(* IEC 61131-3 sources: codesys-ai-industrial-robot-control/plc/src/Comm, 4 files *)

(* ---- GVL_Bridge.st ---- *)
// Exchange with the Python bridge over OPC UA (published by the symbol configuration).
// Tag names for the bridge: config/opcua_tags.yaml. In Phase 1, tests write the inputs.
{attribute 'qualified_only'}
{attribute 'symbol' := 'readwrite'}
VAR_GLOBAL
    // --- inputs (bridge -> PLC) ---
    xHeartbeat : BOOL;                                     // toggled by the bridge every cycle
    xTwinActive : BOOL;                                    // the twin delivers joint feedback
    aJointPosFb : ARRAY[1..6] OF LREAL;                    // measured joint positions [deg]
    aJointTorqueFb : ARRAY[1..6] OF LREAL;                 // measured joint torques [Nm]
    udiFeedbackSeq : UDINT;                                // increments with every feedback sample
    udiFeedbackForSeq : UDINT;                             // udiSetpointSeq the feedback belongs to
    xPE1 : BOOL;                                           // photo-eye at the camera
    xPE2 : BOOL;                                           // photo-eye at the pick window start
    xVacuumOk : BOOL;                                      // vacuum switch of the suction cup
    axBinFull : ARRAY[E_Bin.TypeA..E_Bin.Quarantine] OF BOOL;
    xDoorClosed : BOOL := TRUE;                            // safety door (TRUE = closed)
    xEStopOk : BOOL := TRUE;                               // emergency stop circuit (TRUE = not pressed)
    stVision : ST_VisionMsg;
    stDecision : ST_DecisionMsg;
    xDecisionActive : BOOL;                                // an AI decision service answers stDecision
    // --- outputs (PLC -> bridge) ---
    aJointPosSp : ARRAY[1..6] OF LREAL;                    // joint setpoints [deg]
    udiSetpointSeq : UDINT;                                // increments with every setpoint sample
    lrBeltPos : LREAL;                                     // conveyor position [mm]
    lrBeltVel : LREAL;                                     // conveyor velocity [mm/s]
    xVacuumOn : BOOL;                                      // vacuum valve
    stCapture : ST_CaptureMsg;
    eState : E_PackMLState;
    eMode : E_PackMLMode;
    // --- diagnostics (PLC -> bridge, HMI) ---
    eNewestAlarm : E_AlarmId;
    xAlarmError : BOOL;                                    // an Error-class alarm is active
    xAlarmCritical : BOOL;                                 // a Critical-class alarm is active
    ePickStep : E_PickStep;
    iWorstJoint : INT;                                     // joint with the largest following error
    aFollowingError : ARRAY[1..6] OF LREAL;                // [deg]
END_VAR

(* ---- GVL_Hmi.st ---- *)
// Operator commands from the HMI (CODESYS Visualization) and, for tests and the HMI of later
// phases, over OPC UA (published by the symbol configuration).
{attribute 'qualified_only'}
{attribute 'symbol' := 'readwrite'}
VAR_GLOBAL
    eCommand : E_PackMLCommand;
    eModeRequest : E_PackMLMode := E_PackMLMode.Production;
    xAlarmAck : BOOL;
    axJogPlus : ARRAY[1..6] OF BOOL;
    axJogMinus : ARRAY[1..6] OF BOOL;
    rOverride : REAL := 1.0;                               // speed override ]0, 1]
END_VAR

(* ---- FB_BridgeWatchdog.st ---- *)
(*
    FB_BridgeWatchdog
    Purpose : The Python bridge toggles xHeartbeat every cycle; if it stops toggling for tTimeout
              while enabled, the connection to the digital twin is considered lost.
    Outputs : xLost
    Alarms  : BridgeLost (Critical -> the cell aborts)
*)
FUNCTION_BLOCK FB_BridgeWatchdog
VAR_INPUT
    xHeartbeat : BOOL;
    xEnable : BOOL;
    tTimeout : TIME := T#500MS;
    itfAlarms : I_AlarmSink;
END_VAR
VAR_OUTPUT
    xLost : BOOL;
END_VAR
VAR
    xLastHeartbeat : BOOL;
    tonLost : TON;
END_VAR

tonLost(IN := xEnable AND xHeartbeat = xLastHeartbeat, PT := tTimeout);
xLastHeartbeat := xHeartbeat;
xLost := tonLost.Q;
IF itfAlarms <> 0 THEN
    IF xLost THEN
        itfAlarms.Raise(E_AlarmId.BridgeLost);
    ELSE
        itfAlarms.Clear(E_AlarmId.BridgeLost);
    END_IF
END_IF

(* ---- FB_MessageIntake.st ---- *)
(*
    FB_MessageIntake
    Purpose : Detects new bridge messages by their sequence number, so a message written twice
              (or re-read) is processed only once.
    Outputs : xVisionNew, xDecisionNew - TRUE for one cycle per new message
*)
FUNCTION_BLOCK FB_MessageIntake
VAR_INPUT
    stVision : ST_VisionMsg;
    stDecision : ST_DecisionMsg;
END_VAR
VAR_OUTPUT
    xVisionNew : BOOL;
    xDecisionNew : BOOL;
END_VAR
VAR
    udiLastVisionSeq : UDINT;
    udiLastDecisionSeq : UDINT;
END_VAR

xVisionNew := stVision.udiSeq <> udiLastVisionSeq;
udiLastVisionSeq := stVision.udiSeq;
xDecisionNew := stDecision.udiSeq <> udiLastDecisionSeq;
udiLastDecisionSeq := stDecision.udiSeq;
